(* IEC 61131-3 sources: ironplc/integrations/vscode/src/test/functional/resources, 1 file *)

(* ---- valid.st ---- *)
PROGRAM main
    VAR
        Button AT %IX1: BOOL;
        Buzzer AT %QX1: BOOL;
    END_VAR

    Buzzer := NOT Button;

END_PROGRAM

CONFIGURATION config
    RESOURCE res ON PLC
        TASK plc_task(INTERVAL := T#100ms, PRIORITY := 1);
        PROGRAM plc_task_instance WITH plc_task : main;
    END_RESOURCE
END_CONFIGURATION
